// TwinCAT 3 PLC project PLC1
// ProgramVersion: 3.1.4026.27
// libraries:
//   Tc2_Standard, * (Beckhoff Automation GmbH)
//   Tc2_System, * (Beckhoff Automation GmbH)
// project tree:
//   / PlcTask.TcTTO
//   POUs/ MAIN.TcPOU
// real-time tasks:
//   TASK PlcTask: cycle T#10ms, priority 20, ADS port 350

CONFIGURATION PLC1
    RESOURCE PLC ON TwinCAT3
        TASK PlcTask(INTERVAL := T#10ms, PRIORITY := 20);
        PROGRAM MAIN WITH PlcTask : MAIN;
    END_RESOURCE
END_CONFIGURATION

// ---- POUs/MAIN.TcPOU
PROGRAM MAIN
VAR
    iCount : INT;
    bLight : BOOL;
    bSwitch : BOOL;
END_VAR

iCount := iCount + 1;

// reset logic
IF iCount > 100 THEN
    iCount := 0;
END_IF

// new Light/Switch logic
IF iCount > 50 THEN
    bLight := bSwitch;
ELSE
    bLight := FALSE;
END_IF

END_PROGRAM
